Fanuc KAREL source: ko00075.KL

PROGRAM KO00075
%STACKSIZE=65535
%PRIORITY=65535
%NOLOCKGROUP
VAR
P1 : XYZWPREXT
P2 : XYZWPREXT
F : BOOLEAN
OUT : XYZWPREXT
BEGIN
F=TRUE
-- UNSAFE_SOURCE_IR line 11: OUT = MIRROR(P1, convert_xyzwprext_to_position(P2), F)
END KO00075
